// TIA Portal V19 export
DATA_BLOCK "FctKeyNamePairs"   // DB2000
{ S7_Optimized_Access := 'TRUE'; DB_Accessible_From_OPC_UA := 'FALSE' }
// stored: AutoNumber false, DBAccessibleFromOPCUA false, DBAccessibleFromWebserver false, MemoryReserve 100
   VAR
      VlvL : Array[0..10] of "FctKeyParName";
      PidL { S7_SetPoint := 'True'} : Array[0..10] of "FctKeyParName";
      MotL : Array[0..10] of "FctKeyParName";
      OpAn { S7_SetPoint := 'True'} : Array[0..10] of "FctKeyParName";
   END_VAR
BEGIN
   VlvL[0].Key := 0;
   VlvL[1].Key := 1;
   VlvL[2].Key := 2;
   VlvL[3].Key := 3;
   VlvL[4].Key := 4;
   VlvL[5].Key := 5;
   VlvL[6].Key := 6;
   VlvL[7].Key := 7;
   VlvL[0]."Name" := 'SETLINK';
   VlvL[1]."Name" := 'SETOPR';
   VlvL[2]."Name" := 'SETAUTO';
   VlvL[3]."Name" := 'SETMAN';
   VlvL[4]."Name" := 'SETOPEN';
   VlvL[5]."Name" := 'SETCLOSE';
   VlvL[6]."Name" := 'GETAUTO';
   VlvL[7]."Name" := 'GETOPEN';
   PidL[0].Key := 0;
   PidL[1].Key := 1;
   PidL[2].Key := 2;
   PidL[3].Key := 3;
   PidL[4].Key := 4;
   PidL[5].Key := 5;
   PidL[6].Key := 6;
   PidL[7].Key := 7;
   PidL[0]."Name" := 'SETLINK';
   PidL[1]."Name" := 'SETOPR';
   PidL[2]."Name" := 'SETINT';
   PidL[3]."Name" := 'SETEXT';
   PidL[4]."Name" := 'SETAUTO';
   PidL[5]."Name" := 'SETMAN';
   PidL[6]."Name" := 'SETTRACK';
   PidL[7]."Name" := 'RSTTRACK';
   MotL[0].Key := 0;
   MotL[1].Key := 1;
   MotL[2].Key := 2;
   MotL[3].Key := 3;
   MotL[4].Key := 4;
   MotL[5].Key := 5;
   MotL[6].Key := 6;
   MotL[7].Key := 7;
   MotL[0]."Name" := 'SETLINK';
   MotL[1]."Name" := 'SETOPR';
   MotL[2]."Name" := 'SETAUTO';
   MotL[3]."Name" := 'SETMAN';
   MotL[4]."Name" := 'START';
   MotL[5]."Name" := 'STOP';
   MotL[6]."Name" := 'GETAUTO';
   MotL[7]."Name" := 'STATUS';
   OpAn[0].Key := 0;
   OpAn[1].Key := 1;
   OpAn[2].Key := 2;
   OpAn[3].Key := 3;
   OpAn[4].Key := 4;
   OpAn[5].Key := 5;
   OpAn[0]."Name" := 'SETLINK';
   OpAn[1]."Name" := 'SETOPR';
   OpAn[2]."Name" := 'SETINT';
   OpAn[3]."Name" := 'SETEXT';
   OpAn[4]."Name" := 'SETOPEN';
   OpAn[5]."Name" := 'SETCLOSE';
END_DATA_BLOCK
